//{attribute 'qualified_only'}
VAR_GLOBAL CONSTANT
	//C_Max_ErrorList				: INT:=200;
	//C_Max_Pistons				: INT:=7;
	//C_Max_MotorsAC				: INT:=6;
	//C_Max_Measure				: INT:=15;
END_VAR

(* stored: Version 1.1.0.1, ProductVersion 3.1.4024.13
   GVL Global_Constant: Id {77daaa20-5a1d-486c-b8b4-df6b9b3f5848} *)
